RoboDK station: PICK2.rdk

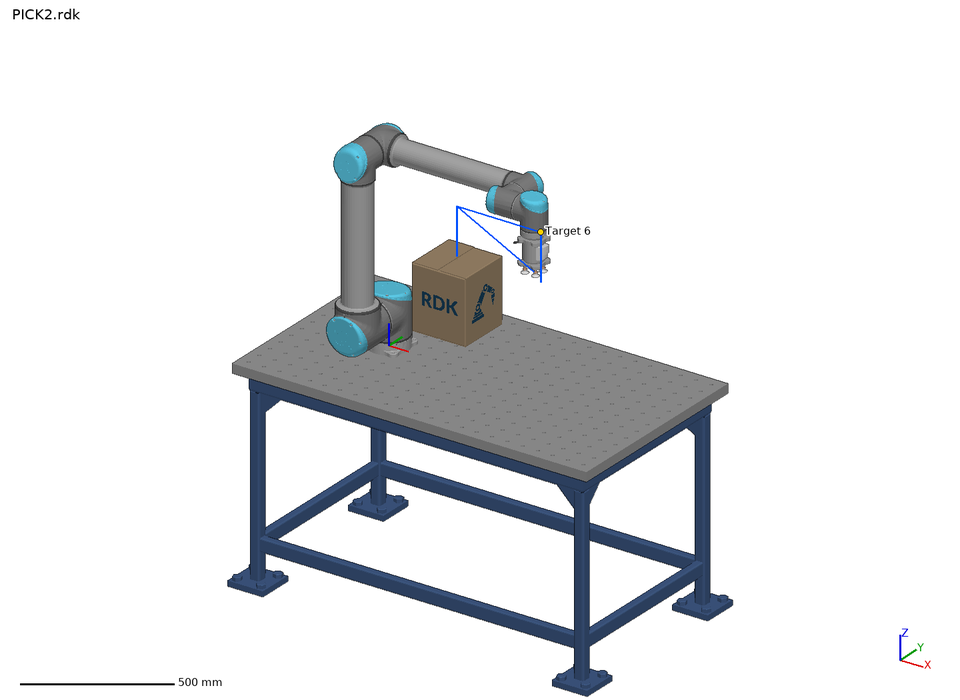
[picture v0: the station drawn from its stored meshes, robots at their saved joint values, targets as dots, program paths as lines]
Station PICK2 (saved by RoboDK 6.1.1). Poses are relative to the parent item; angles as X-Y-Z fixed-axis rotations.
  - frame UR10 Base at (0, 0, 0) mm
    - robot UR10: 6 axes, payload 10 kg, reach 1300 mm, repeatability 0.1 mm, weight 28.9 kg
        modified DH rows (alpha deg, a mm, theta deg, d mm): 0, 0, 0, 128; 90, 0, 180, 0; 0, 612.7, 0, 0; 0, 571.6, 0, 163.9; -90, 0, 0, 115.7; 90, 0, 180, 92.2
        joint limits [-360, -360, -360, -360, -360, -360] to [360, 360, 360, 360, 360, 360]; home [0, -90, -90, 0, 90, 0]; saved at [0, -90, -90, -90, 90, 0]
      - tool SMC ZXP7A01-ZP25C-X1 Vacuum Gripper, TCP at (0, 0, 125) mm, size 88 x 106.8 x 127.9 mm
    - target Target 6 (Cartesian target) at (436.45, 233.38, 436.43) mm, rotated rx 180 ry 0 rz 0 deg; joints [0, -90, -90, -90, 90, 0] of UR10
    - object Box 215x215mm (Folded) at (0, 130, 124.22) mm, size 213.4 x 213.4 x 248.4 mm, geometry from Box-215x215mm-Folded.sld
  - object Table 1400x800x800mm at (0, 0, 0) mm, size 1420 x 820 x 800 mm, geometry from Table-1400x800x800mm.sld
  - Python program Prog1 (listed below)
  - program PickPlace_UR10_IDA_VUELTA (20 instructions, listed below)
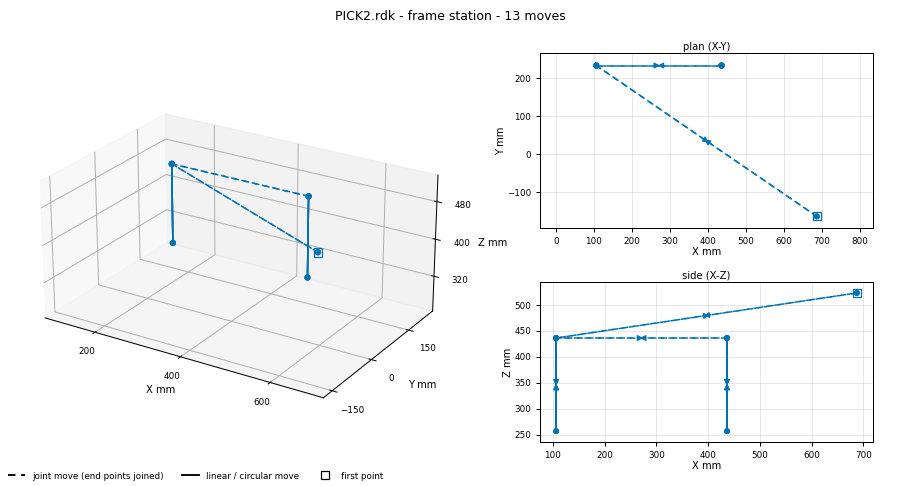
[picture p0: tool path of PICK2.rdk in frame station, 13 of 13 moves have a stored position in this frame; points joined in program order, loops and branches not executed]

--- Python program Prog1 ---
# -*- coding: utf-8 -*-
"""
PICK & PLACE UR10 + pinza SMC en RoboDK - DESDE CERO.

Estacion necesaria (NO hace falta ningun target previo):
    UR10
    SMC ZXP7A01... (herramienta hija del UR10)
    Table 1400x800x800mm
    Box 215x215mm (Folded)

Al ejecutar Prog1:
  1) Recoloca la caja dentro de la mesa.
  2) CREA home, aprox1, pick, aprox2, place, Target 6.
  3) CREA PickPlace_UR10_IDA_VUELTA.
  4) SIMULA tomar la caja, moverla, devolverla y regresar a home.

Se usa exclusivamente el SIMULADOR. No activa succion real.
Guarda una copia de la estacion antes de ejecutarlo.
"""

import json
import math
from robodk.robolink import *
from robodk.robomath import *

# =============== PERSONALIZA SOLO SI HACE FALTA ===============
HOME_ARTICULACIONES = [0, -90, -90, -90, 90, 0]  # Grados
MARGEN_BORDE_MM = 35            # Caja separada del borde de la mesa
SEPARACION_BASE_MM = 225        # Evitar colocar caja pegada a la base
SUBIDA_SEGURA_MM = 180         # Aproximaciones por encima de la caja
HOLGURA_TCP_MM = 8             # TCP unos mm por ENCIMA de la tapa, no de la mesa
DISTANCIA_TRASLADO_MM = 330
VELOCIDAD_LINEAL_MM_S = 80
VELOCIDAD_SIMULACION = 1.0      # 1.0 = velocidad de simulacion normal
AUTO_EJECUTAR = True           # True: anima al ejecutar Prog1 por primera vez
MOSTRAR_FLECHAS_TARGETS = False
NOMBRE_PROGRAMA = 'PickPlace_UR10_IDA_VUELTA'
# ==============================================================

RDK = Robolink()
RDK.setRunMode(RUNMODE_SIMULATE)  # Solo simulacion, NUNCA el robot real


def buscar_objeto(prefijo):
    for elemento in RDK.ItemList(ITEM_TYPE_OBJECT):
        if elemento.Name().lower().startswith(prefijo.lower()):
            return elemento
    raise Exception('Falta el objeto llamado: ' + prefijo)


def limites_mundo(elemento):
    """BoundingBox de RoboDK: coordenadas globales (mm)."""
    datos = elemento.setParam('BoundingBox')
    if isinstance(datos, str):
        datos = json.loads(datos)
    if not isinstance(datos, dict):
        raise Exception('No puedo medir la geometria de ' + elemento.Name())
    datos = {str(k).lower(): v for k, v in datos.items()}
    minimo = datos.get('min', datos.get('xyzmin'))
    maximo = datos.get('max', datos.get('xyzmax'))
    if minimo is None or maximo is None:
        raise Exception('BoundingBox inesperado en ' + elemento.Name() + ': ' + str(datos))
    return [float(v) for v in minimo[:3]], [float(v) for v in maximo[:3]]


def limitar(v, menor, mayor):
    return max(menor, min(mayor, v))


# =========== 1. ENCONTRAR LOS OBJETOS YA IMPORTADOS ===========
robot = RDK.Item('UR10', ITEM_TYPE_ROBOT)
if not robot.Valid():
    raise Exception('No se encuentra UR10. Importa primero el robot.')

pinzas = [e for e in robot.Childs() if e.Type() == ITEM_TYPE_TOOL]
if not pinzas:
    pinza_vinculada = robot.getLink(ITEM_TYPE_TOOL)
    if pinza_vinculada.Valid():
        pinzas = [pinza_vinculada]
if not pinzas:
    raise Exception('No encuentro la herramienta SMC debajo del UR10.')
pinza = pinzas[0]

mesa = buscar_objeto('Table 1400x800')
caja = buscar_objeto('Box 215x215')

# La referencia en la estacion mostrada es UR10 Base.
referencia = robot.Parent()
if referencia.Type() != ITEM_TYPE_FRAME:
    referencia = robot.getLink(ITEM_TYPE_FRAME)
if not referencia.Valid():
    raise Exception('No encuentro UR10 Base.')

# Si la caja se quedo agarrada tras otra simulacion, la soltamos
# conservando su posicion absoluta antes de medirla.
caja.setParentStatic(referencia)
robot.setPoseFrame(referencia)
robot.setPoseTool(pinza)

# =========== 2. MEDIR LA MESA Y LA CAJA ===========
mesa_min, mesa_max = limites_mundo(mesa)
caja_min, caja_max = limites_mundo(caja)

ancho_caja = caja_max[0] - caja_min[0]
largo_caja = caja_max[1] - caja_min[1]
alto_caja = caja_max[2] - caja_min[2]
superficie_mesa = mesa_max[2]

if min(ancho_caja, largo_caja, alto_caja) <= 1:
    raise Exception('La caja tiene dimensiones invalidas. Revisa el modelo.')

# El CENTRO de la caja debe dejar margen para TODA la caja.
x_min = mesa_min[0] + MARGEN_BORDE_MM + ancho_caja / 2.0
x_max = mesa_max[0] - MARGEN_BORDE_MM - ancho_caja / 2.0
y_min = mesa_min[1] + MARGEN_BORDE_MM + largo_caja / 2.0
y_max = mesa_max[1] - MARGEN_BORDE_MM - largo_caja / 2.0
if x_min >= x_max or y_min >= y_max:
    raise Exception('La caja no cabe en la zona util de la mesa.')

x_original = limitar((caja_min[0] + caja_max[0]) / 2.0, x_min, x_max)
y_original = limitar((caja_min[1] + caja_max[1]) / 2.0, y_min, y_max)

base_robot = robot.PoseAbs().Pos()


def alejado_de_base(x, y):
    return math.hypot(x - base_robot[0], y - base_robot[1]) >= SEPARACION_BASE_MM


# La pinza siempre apunta verticalmente hacia la caja.
# Las poses de los objetivos se guardan relativas a UR10 Base.
mundo_a_referencia = referencia.PoseAbs().inv()
pose_herramienta = robot.PoseTool()
pose_referencia = robot.PoseFrame()


def pose_objetivo(x, y, z, rotacion):
    pose_absoluta = transl(x, y, z) * rotz(rotacion) * rotx(math.pi)
    return mundo_a_referencia * pose_absoluta


def se_alcanza(pose):
    try:
        articulaciones = robot.SolveIK(
            pose, HOME_ARTICULACIONES, pose_herramienta, pose_referencia)
        return len(articulaciones.list()) >= 6
    except Exception:
        return False


# El TCP NO debe llegar al tablero: PICK/PLACE quedan a la altura de la
# TAPA DE LA CAJA, con algunos mm adicionales de holgura.
z_pick = superficie_mesa + alto_caja + HOLGURA_TCP_MM
z_aprox = z_pick + SUBIDA_SEGURA_MM

# Para conservar el comportamiento del PRIMER codigo que ya te funciono,
# usamos las mismas alternativas para encontrar un recorrido alcanzable.
origines = [(x_original, y_original)]
for dx, dy in [(0, 130), (0, -130), (-150, 0), (150, 0),
               (-230, 120), (-230, -120), (230, 120), (230, -120)]:
    candidato = (limitar(x_original + dx, x_min, x_max),
                 limitar(y_original + dy, y_min, y_max))
    if candidato not in origines:
        origines.append(candidato)

traslados = [
    (DISTANCIA_TRASLADO_MM, 0), (-DISTANCIA_TRASLADO_MM, 0),
    (0, DISTANCIA_TRASLADO_MM), (0, -DISTANCIA_TRASLADO_MM),
    (280, 180), (280, -180), (-280, 180), (-280, -180),
    (250, 0), (-250, 0), (0, 250), (0, -250)
]

solucion = None
for giro in [0, math.pi / 2, math.pi, -math.pi / 2]:
    for xp, yp in origines:
        if not alejado_de_base(xp, yp):
            continue
        p_pick = pose_objetivo(xp, yp, z_pick, giro)
        p_aprox1 = pose_objetivo(xp, yp, z_aprox, giro)
        if not (se_alcanza(p_pick) and se_alcanza(p_aprox1)):
            continue

        for dx, dy in traslados:
            x_destino, y_destino = xp + dx, yp + dy
            if not (x_min <= x_destino <= x_max and
                    y_min <= y_destino <= y_max):
                continue
            if not alejado_de_base(x_destino, y_destino):
                continue
            if math.hypot(dx, dy) <= max(ancho_caja, largo_caja) + 30:
                continue
            p_place = pose_objetivo(x_destino, y_destino, z_pick, giro)
            p_aprox2 = pose_objetivo(x_destino, y_destino, z_aprox, giro)
            if se_alcanza(p_place) and se_alcanza(p_aprox2):
                solucion = (xp, yp, x_destino, y_destino,
                            p_pick, p_aprox1, p_place, p_aprox2)
                break
        if solucion is not None:
            break
    if solucion is not None:
        break

if solucion is None:
    raise Exception(
        'No se encontraron dos puntos alcanzables dentro de la mesa. '
        'Comprueba la posicion de la mesa, la pinza y su TCP.')

xp, yp, xd, yd, p_pick, p_aprox1, p_place, p_aprox2 = solucion

# =========== 3. RECOLOCAR LA CAJA EN SU ORIGEN ===========
# Recolocacion antes de generar el programa. Asi, si ejecutas Prog1 otra
# vez, no se queda la caja donde termino la simulacion anterior.
centro_caja_x = (caja_min[0] + caja_max[0]) / 2.0
centro_caja_y = (caja_min[1] + caja_max[1]) / 2.0
caja.setPoseAbs(
    transl(xp - centro_caja_x,
           yp - centro_caja_y,
           superficie_mesa - caja_min[2]) * caja.PoseAbs())

# =========== 4. CREAR TODOS LOS TARGETS DESDE CERO ===========
# Es importante eliminar primero el programa que los utiliza.
programa_viejo = RDK.Item(NOMBRE_PROGRAMA, ITEM_TYPE_PROGRAM)
if programa_viejo.Valid():
    programa_viejo.Delete()

for nombre in ['home', 'aprox1', 'pick', 'aprox2', 'place', 'Target 6']:
    anterior = RDK.Item(nombre, ITEM_TYPE_TARGET)
    if anterior.Valid():
        anterior.Delete()


def crear_cartesiano(nombre, pose):
    objetivo = RDK.AddTarget(nombre, referencia, robot)
    objetivo.setAsCartesianTarget()
    objetivo.setPose(pose)
    objetivo.setVisible(MOSTRAR_FLECHAS_TARGETS)
    return objetivo


home = RDK.AddTarget('home', referencia, robot)
home.setAsJointTarget()
home.setJoints(HOME_ARTICULACIONES)
home.setVisible(MOSTRAR_FLECHAS_TARGETS)

aprox1 = crear_cartesiano('aprox1', p_aprox1)
pick = crear_cartesiano('pick', p_pick)
aprox2 = crear_cartesiano('aprox2', p_aprox2)
place = crear_cartesiano('place', p_place)
retirada = crear_cartesiano('Target 6', p_aprox2)

# =========== 5. CREAR PROGRAMA DE IDA Y VUELTA ===========
prog = RDK.AddProgram(NOMBRE_PROGRAMA, robot)
prog.setPoseFrame(referencia)
prog.setPoseTool(pinza)
prog.setSpeed(VELOCIDAD_LINEAL_MM_S)
prog.setRunType(PROGRAM_RUN_ON_SIMULATOR)


def tomar_caja(nombre_evento):
    # El MISMO formato de evento del primer script que ya funcionaba.
    prog.setParam('Add', {
        'Name': nombre_evento,
        'Type': 7,
        'Behavior': 0,
        'ToolPtr': str(pinza.item),
        'ObjectList': str(caja.item),
        'AttachStrategy': 4,
        'AttachDistance': 200
    })


def soltar_caja(nombre_evento):
    prog.setParam('Add', {
        'Name': nombre_evento,
        'Type': 7,
        'Behavior': 1,
        'ToolPtr': str(pinza.item),
        'FramePtr': str(referencia.item)
    })


# IDA: original -> segundo lugar
prog.MoveJ(home)
prog.MoveJ(aprox1)
prog.MoveL(pick)
tomar_caja('1 - Tomar caja en PICK')
prog.MoveL(aprox1)
prog.MoveJ(aprox2)
prog.MoveL(place)
soltar_caja('2 - Soltar caja en PLACE')
prog.MoveL(aprox2)

# VUELTA: segundo lugar -> original
prog.MoveL(place)
tomar_caja('3 - Tomar caja en PLACE')
prog.MoveL(aprox2)
prog.MoveJ(aprox1)
prog.MoveL(pick)
soltar_caja('4 - Devolver caja a PICK')
prog.MoveL(aprox1)
prog.MoveJ(home)

prog.ShowInstructions(True)
prog.ShowTargets(MOSTRAR_FLECHAS_TARGETS)

print('OK. Se crearon: home, aprox1, pick, aprox2, place y Target 6.')
print('OK. Programa creado: ' + NOMBRE_PROGRAMA)
print('CAJA INICIAL: X=%.1f Y=%.1f mm' % (xp, yp))
print('CAJA DESTINO: X=%.1f Y=%.1f mm' % (xd, yd))
print('Altura de mesa=%.1f; altura de caja=%.1f; TCP de pick=%.1f mm' %
      (superficie_mesa, alto_caja, z_pick))
print('Secuencia: tomar, colocar, volver a tomar y devolver al origen.')

# =========== 6. INICIAR SIMULACION EN PRIMERA EJECUCION ===========
# Sin prog.Update(): la version anterior se bloqueaba al validar un programa
# antes de simularlo. Si RoboDK no puede iniciarlo, queda creado en el arbol.
if AUTO_EJECUTAR:
    try:
        RDK.setRunMode(RUNMODE_SIMULATE)
        RDK.setSimulationSpeed(VELOCIDAD_SIMULACION)
        resultado = prog.RunCode()
        if resultado <= 0:
            print('AVISO: El programa existe pero RoboDK no inicio la animacion.')
            print('Abre el programa del arbol y revisa que sus movimientos sean validos.')
        else:
            print('SIMULACION INICIADA. No necesitas hacer doble clic.')
    except Exception as error:
        print('AVISO: No se inicio automaticamente: ' + str(error))
        print('El programa SI esta creado. Haz doble clic en ' + NOMBRE_PROGRAMA)
else:
    print('Para simular, haz doble clic en ' + NOMBRE_PROGRAMA)

print('IMPORTANTE: Simulacion solamente. Revisar TCP y colisiones antes de usar un robot real.')

--- program PickPlace_UR10_IDA_VUELTA (robot UR10) ---
  Est. Ref.: UR10 Base
  Est. herr: SMC ZXP7A01-ZP25C-X1 Vacuum Gripper
  Establecer velocidad (80.0 mm/s)
  MoveJ (home) to (687.3, -163.9, 523.5) mm, rotated rx -180 ry 0 rz -90 deg; joints [0, -90, -90, -90, 90, 0]
  MoveJ (aprox1) to (106.45, 233.38, 436.43) mm, rotated rx 180 ry 0 rz 0 deg; joints [0, -90, -90, -90, 90, 0]
  MoveL (pick) to (106.45, 233.38, 256.43) mm, rotated rx 180 ry 0 rz 0 deg; joints [0, -90, -90, -90, 90, 0]
  1 - Tomar caja en PICK
  MoveL (aprox1) to (106.45, 233.38, 436.43) mm, rotated rx 180 ry 0 rz 0 deg; joints [0, -90, -90, -90, 90, 0]
  MoveJ (aprox2) to (436.45, 233.38, 436.43) mm, rotated rx 180 ry 0 rz 0 deg; joints [0, -90, -90, -90, 90, 0]
  MoveL (place) to (436.45, 233.38, 256.43) mm, rotated rx 180 ry 0 rz 0 deg; joints [0, -90, -90, -90, 90, 0]
  2 - Soltar caja en PLACE
  MoveL (aprox2) to (436.45, 233.38, 436.43) mm, rotated rx 180 ry 0 rz 0 deg; joints [0, -90, -90, -90, 90, 0]
  MoveL (place) to (436.45, 233.38, 256.43) mm, rotated rx 180 ry 0 rz 0 deg; joints [0, -90, -90, -90, 90, 0]
  3 - Tomar caja en PLACE
  MoveL (aprox2) to (436.45, 233.38, 436.43) mm, rotated rx 180 ry 0 rz 0 deg; joints [0, -90, -90, -90, 90, 0]
  MoveJ (aprox1) to (106.45, 233.38, 436.43) mm, rotated rx 180 ry 0 rz 0 deg; joints [0, -90, -90, -90, 90, 0]
  MoveL (pick) to (106.45, 233.38, 256.43) mm, rotated rx 180 ry 0 rz 0 deg; joints [0, -90, -90, -90, 90, 0]
  4 - Devolver caja a PICK
  MoveL (aprox1) to (106.45, 233.38, 436.43) mm, rotated rx 180 ry 0 rz 0 deg; joints [0, -90, -90, -90, 90, 0]
  MoveJ (home) to (687.3, -163.9, 523.5) mm, rotated rx -180 ry 0 rz -90 deg; joints [0, -90, -90, -90, 90, 0]
